// TIA Portal V20 export
ORGANIZATION_BLOCK "T7_OB30"   // OB30, LAD, CyclicInterrupt
TITLE = T7_OB30
{ S7_Optimized_Access := 'TRUE' }
AUTHOR : IA
FAMILY : PRUEBA
VERSION : 0.1
// Tanda 3: CyclicInterrupt, incrementa OB30_Cuenta
// stored: AutoNumber false, IsIECCheckEnabled false, SetENOAutomatically false
   VAR_INPUT
      Initial_Call : Bool;
      Event_Count : Int;
   END_VAR
BEGIN

REGION Network 1: Contador de vida
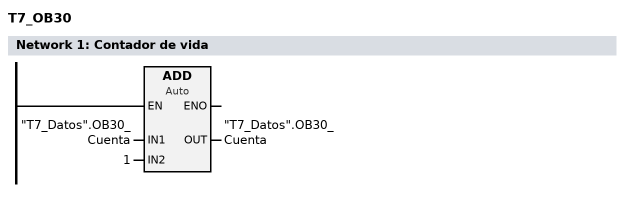
   RUNG wire#powerrail
      Add(in1 := "T7_Datos".OB30_Cuenta, in2 := 1, out => "T7_Datos".OB30_Cuenta)
   END_RUNG
   // the same network as SCL:
   "T7_Datos".OB30_Cuenta := "T7_Datos".OB30_Cuenta + 1;
END_REGION
END_ORGANIZATION_BLOCK
